SUBAPPLICATION Uebung_OPC_L08_AX (* Wie Training_08, lokal: SoftKey_F1 ruft die Toggle-Methode per localhost auf, Flipflop schaltet Output_Q1 *)
  (* Standard: 61499-2; Description: Copyright (c) 2026 Meisterschulen am Ostbahnhof This program and the accompanying materials are made available under the terms of the Eclipse Public License 2.0 which is available at https://www.eclipse.org/legal/epl-2.0/ SPDX-License-Identifier: EPL-2.0 *)
  (* Version 1.0, 2026-10-18, Franz Höpfinger, Meisterschulen am Ostbahnhof, Aus SubApp_PC_A + SubApp_PC_B von test_VV zusammengefuehrt, lokale Varianten der Bausteine *)
  PACKAGE Meins::OPC_UA_Lokal;
  IMPORT Uebungen::const::UT::DefaultPool::SoftKey_F1;
  IMPORT Meins::OPC_UA_Lokal::const::OpcUaLokal::FF1_TRIGGER_CALL;
  IMPORT Meins::OPC_UA_Lokal::const::OpcUaLokal::FF1_STATE_READ;
  IMPORT logiBUS::io::DQ::logiBUS_DO::Output_Q1;
  IMPORT Meins::OPC_UA_Lokal::const::OpcUaLokal::FF1_TRIGGER_METHOD;
  IMPORT Meins::OPC_UA_Lokal::const::OpcUaLokal::FF1_STATE_WRITE;
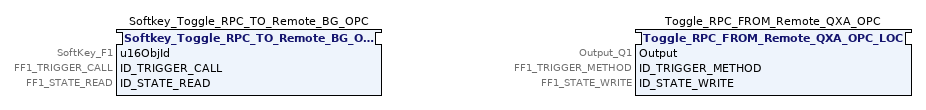
  SUBAPPS
    Softkey_Toggle_RPC_TO_Remote_BG_OPC : MyLib::sys::Softkey_Toggle_RPC_TO_Remote_BG_OPC(u16ObjId := SoftKey_F1, ID_TRIGGER_CALL := FF1_TRIGGER_CALL, ID_STATE_READ := FF1_STATE_READ);
    Toggle_RPC_FROM_Remote_QXA_OPC : MyLib::sys::Toggle_RPC_FROM_Remote_QXA_OPC_LOC(Output := Output_Q1, ID_TRIGGER_METHOD := FF1_TRIGGER_METHOD, ID_STATE_WRITE := FF1_STATE_WRITE);
  END_SUBAPPS
END_SUBAPPLICATION
